Fanuc KAREL source: ka00145.KL

PROGRAM KA00145
%STACKSIZE=65535
%PRIORITY=65535
%NOLOCKGROUP
VAR
SRC : ARRAY[4] OF INTEGER
DST : ARRAY[4] OF INTEGER
BEGIN
-- UNRESOLVED_PC line 7 opcodes [22 22 1E] marker_code=0
END KA00145
